# EPICS substitutions: iocBoot/iocTomoScan_19BM/tomoScan.substitutions
# Edited by ALK 10/23/2026 to match current beamline configuration.
#
#
# SAMPLE_X and SAMPLE_Y are the hexapod's X and Y axes.
#     m1 Hexapod X  mm   +/-27.5      m4 Hexapod A  deg  +/-7.5
#     m2 Hexapod Y  mm   +/-30        m5 Hexapod B  deg  +/-7.5
#     m3 Hexapod Z  mm   0+/-27.5     m6 Hexapod C  deg  +/-15
#
# SAMPLE_X / SAMPLE_Y are the translations UNDER the rotary, which tomoscan
# uses to move the sample clear of the beam for flat fields.  They are NOT the
# SampleTop X/Z pair on top of the rotary -- a Kohzu CYAT-070 stage which co-rotates with
# theta and centres the sample on the rotation axis.  That pair is set by hand
# and has no tomoscan binding; do not rebind these macros to it once it is
# wired.
#
# The hexapod runs on an Aerotech Automation1,  a different
# controller from the Ensemble that drives the rotation, so 19-BM will end up
# with two Aerotech controllers (actually, three including the controller for
# Optics_Z, but TomoScan doesn't need to know about that).
#
# ROTATION is 19bmSoft:aero:m1, confirmed by the beamline 2026-09-19.  It is the
# Aerotech Ensemble air-bearing rotary stage, served by the 19bmSoft IOC on
# hounsfield.
#
# CAMERA is the bare areaDetector IOC prefix; tomoscan.py appends "cam1:" itself.
# The 19-BM camera is a Vieworks VP-61MX (9568x6380, UInt16) on a Euresys
# Coaxlink grabber, driven by ADEuresys via ADGenICam.  Its IOC lives in
# /net/s19dserv/xorApps/epics/synApps_6_3/ioc/19bmVieworks and loads the
# standard commonPlugins.cmd set, so HDF1:, Pva1:, ROI1: and CB1: all exist.
file "$(TOP)/db/tomoScan.template"
{
pattern
{  P,       R,           CAMERA,          FILE_PLUGIN,          ROTATION,        SAMPLE_X,        SAMPLE_Y,           CLOSE_SHUTTER,        CLOSE_VALUE,          OPEN_SHUTTER,         OPEN_VALUE}
{19bm:, TomoScan:, 19bmVieworks:, 19bmVieworks:HDF1:, 19bmSoft:aero:m1, 19bmHXP:m1, 19bmHXP:m2, S19BM-PSS:FES:CloseEPICSC,       1,       S19BM-PSS:FES:OpenEPICSC,       1}
}

# For the Ensemble PSO_ENC_PER_ROTATION is a signed number containing the number of encoder pulses per rotation in positive dial coordinates
#
# These four values are NOT placeholders.  19-BM inherits the rotary stage and
# its Aerotech Ensemble controller from 7-BM intact, and all four are
# properties of that hardware rather than of where it is plugged in, so they
# carry over unchanged from iocTomoScan_7BM/tomoScan.substitutions.
#
# PSO_ENC_PER_ROTATION is positive at 19-BM: after remounting, the encoder
# counts increase as the dial position increases (confirmed 2026-10-23, opposite
# of the 7-BM wiring this stage came from).  If the stage is ever remounted
# again, re-verify the SIGN the way 32-ID-C documents: compare the signs of
# the rotation motor's .RVAL and .DRBV, which must agree for a positive value.
file "$(TOP)/db/tomoScan_PSO.template"
{
pattern
{  P,       R,      PSO_MODEL, PSO_PORT, PSO_AXIS_NAME, PSO_ENC_INPUT, PSO_ENC_PER_ROTATION}
{19bm:, TomoScan:,      0,     PSO_PORT,       A,             3,             8192000.}
}

# Beamline-specific template.  Modeled on 7-BM rather than 32-ID-C because
# 32-ID-C's template carries an mctOptics prefix that 19-BM has no server for;
# the optics metadata records live in tomoScan_19BM.template itself.
#
# LINE is the GenICam TriggerSource the PSO output is wired to.  The Vieworks
# VP-61MX offers Software, UserOutput0, LinkTrigger0, Timer0Active and Line0.
# 19-BM has only the front-end shutter, bound through OPEN_SHUTTER /
# CLOSE_SHUTTER above; there are no fast-shutter macros because
# tomoScan_19BM.template defines no fast-shutter records.
#
# SHUTTER_STATUS reports whether the beam is BLOCKED: 1 = closed, 0 = open.
# That is the inverse of the PA:...:STA_?_SBS_OPEN_PL records used at 32-ID,
# and matches what 2-BM-B does with S02BM-PSS:SBS:BeamBlockingM.  The .VAL
# suffix follows 2-BM-B.
#
# BEAM_READY mirrors 2-BM-B, which uses S02BM-PSS:FES:FEEPSPermitM.
file "$(TOP)/db/tomoScan_19BM.template"
{
pattern
{  P,       R,             BEAM_READY,        READY_VALUE,          SHUTTER_STATUS,           LINE}
{19bm:, TomoScan:, S19BM-PSS:FES:FEEPSPermitM,      1,      S19BM-PSS:FES:BeamBlockingM.VAL, Line0}
}
